Fanuc KAREL source: KT00241.KL

PROGRAM KT00241
%NOLOCKGROUP
VAR
  Y1: ARRAY[2] OF BYTE
  B2: BOOLEAN
  OUT: BOOLEAN
BEGIN
  Y1[1] = 2
    B2 = FALSE
  OUT = Y1[1] OR B2
END KT00241
